(* IEC 61131-3 sources: plc-st-coding-agent/progress/evidence/f14_v5_public_pilot_20261112/jobs/custom_minimax-m27, 20 files *)

(* ---- public-easy-01.candidate_01.st ---- *)
FUNCTION_BLOCK FillingLineControl
VAR_INPUT
    bottleSensor          : BOOL;
    cleaningConfirmButton : BOOL;
    fillingConfirmButton  : BOOL;
    cappingConfirmButton  : BOOL;
    packingConfirmButton  : BOOL;
    finishedButton        : BOOL;
END_VAR
VAR_OUTPUT
    Pump_Motor       : BOOL;
    Filling_Valve    : BOOL;
    Capping_Machine  : BOOL;
    Packing_Machine  : BOOL;
    Completion_Light : BOOL;
END_VAR
VAR
    eState : INT;
END_VAR

// ENGINEERING_CONTRACT
// States: 0=IDLE, 1=CLEANING, 2=FILLING, 3=CAPPING, 4=PACKING, 5=COMPLETED
// PUB003: bottleSensor triggers pump motor continuously (retriggers if bottle stays)
// PUB004-PUB007: Each confirm button advances to next stage; next output activates immediately
// PUB008: finishedButton resets to IDLE; all outputs deactivate, Completion_Light clears
// Output retention: No output holds state beyond its stage; Completion_Light is latched until reset
// Same-scan priority: Transition logic evaluated after output assignments per state
// Boundaries: bottleSensor edge-sensitive to detected; confirm buttons level-triggered per stage

CASE eState OF
    0: // IDLE
        Pump_Motor       := FALSE;
        Filling_Valve    := FALSE;
        Capping_Machine  := FALSE;
        Packing_Machine  := FALSE;
        Completion_Light := FALSE;
        IF bottleSensor THEN
            eState := 1;
        END_IF;

    1: // CLEANING
        Pump_Motor       := TRUE;
        Filling_Valve    := FALSE;
        Capping_Machine  := FALSE;
        Packing_Machine  := FALSE;
        Completion_Light := FALSE;
        IF cleaningConfirmButton THEN
            eState := 2;
        END_IF;

    2: // FILLING
        Pump_Motor       := FALSE;
        Filling_Valve    := TRUE;
        Capping_Machine  := FALSE;
        Packing_Machine  := FALSE;
        Completion_Light := FALSE;
        IF fillingConfirmButton THEN
            eState := 3;
        END_IF;

    3: // CAPPING
        Pump_Motor       := FALSE;
        Filling_Valve    := FALSE;
        Capping_Machine  := TRUE;
        Packing_Machine  := FALSE;
        Completion_Light := FALSE;
        IF cappingConfirmButton THEN
            eState := 4;
        END_IF;

    4: // PACKING
        Pump_Motor       := FALSE;
        Filling_Valve    := FALSE;
        Capping_Machine  := FALSE;
        Packing_Machine  := TRUE;
        Completion_Light := FALSE;
        IF packingConfirmButton THEN
            eState := 5;
        END_IF;

    5: // COMPLETED
        Pump_Motor       := FALSE;
        Filling_Valve    := FALSE;
        Capping_Machine  := FALSE;
        Packing_Machine  := FALSE;
        Completion_Light := TRUE;
        IF finishedButton THEN
            eState := 0;
        END_IF;

END_CASE;

END_FUNCTION_BLOCK

(* ---- public-easy-01.candidate_02.st ---- *)
FUNCTION_BLOCK FillingLineControl
VAR_INPUT
    bottleSensor          : BOOL;
    cleaningConfirmButton : BOOL;
    fillingConfirmButton  : BOOL;
    cappingConfirmButton  : BOOL;
    packingConfirmButton  : BOOL;
    finishedButton        : BOOL;
END_VAR
VAR_OUTPUT
    Pump_Motor       : BOOL;
    Filling_Valve    : BOOL;
    Capping_Machine  : BOOL;
    Packing_Machine  : BOOL;
    Completion_Light : BOOL;
END_VAR
VAR
    eState    : INT;
    nextState : INT;
END_VAR

// ENGINEERING_CONTRACT
// States: 0=IDLE, 1=CLEANING, 2=FILLING, 3=CAPPING, 4=PACKING, 5=COMPLETED
// PUB003: bottleSensor triggers pump motor continuously (retriggers if bottle stays)
// PUB004-PUB007: Each confirm button advances to next stage; next output activates immediately
// PUB008: finishedButton resets to IDLE; all outputs deactivate, Completion_Light clears
// Output retention: No output holds state beyond its stage; Completion_Light is latched until reset
// Same-scan priority: Two-CASE pattern prevents premature output assignment during transition evaluation
// Boundaries: bottleSensor edge-sensitive to detected; confirm buttons level-triggered per stage

nextState := eState;
CASE eState OF
    0:
        IF bottleSensor THEN
            nextState := 1;
        END_IF;
    1:
        IF cleaningConfirmButton THEN
            nextState := 2;
        END_IF;
    2:
        IF fillingConfirmButton THEN
            nextState := 3;
        END_IF;
    3:
        IF cappingConfirmButton THEN
            nextState := 4;
        END_IF;
    4:
        IF packingConfirmButton THEN
            nextState := 5;
        END_IF;
    5:
        IF finishedButton THEN
            nextState := 0;
        END_IF;
END_CASE;

eState := nextState;

CASE eState OF
    0:
        Pump_Motor       := FALSE;
        Filling_Valve    := FALSE;
        Capping_Machine  := FALSE;
        Packing_Machine  := FALSE;
        Completion_Light := FALSE;
    1:
        Pump_Motor       := TRUE;
        Filling_Valve    := FALSE;
        Capping_Machine  := FALSE;
        Packing_Machine  := FALSE;
        Completion_Light := FALSE;
    2:
        Pump_Motor       := FALSE;
        Filling_Valve    := TRUE;
        Capping_Machine  := FALSE;
        Packing_Machine  := FALSE;
        Completion_Light := FALSE;
    3:
        Pump_Motor       := FALSE;
        Filling_Valve    := FALSE;
        Capping_Machine  := TRUE;
        Packing_Machine  := FALSE;
        Completion_Light := FALSE;
    4:
        Pump_Motor       := FALSE;
        Filling_Valve    := FALSE;
        Capping_Machine  := FALSE;
        Packing_Machine  := TRUE;
        Completion_Light := FALSE;
    5:
        Pump_Motor       := FALSE;
        Filling_Valve    := FALSE;
        Capping_Machine  := FALSE;
        Packing_Machine  := FALSE;
        Completion_Light := TRUE;
END_CASE;

END_FUNCTION_BLOCK

(* ---- public-easy-01.raw_candidate_01.st ---- *)
FUNCTION_BLOCK FillingLineControl
VAR_INPUT
    bottleSensor          : BOOL;
    cleaningConfirmButton : BOOL;
    fillingConfirmButton  : BOOL;
    cappingConfirmButton  : BOOL;
    packingConfirmButton  : BOOL;
    finishedButton        : BOOL;
END_VAR
VAR_OUTPUT
    Pump_Motor       : BOOL;
    Filling_Valve    : BOOL;
    Capping_Machine  : BOOL;
    Packing_Machine  : BOOL;
    Completion_Light : BOOL;
END_VAR
VAR
    eState : INT;
END_VAR

// ENGINEERING_CONTRACT
// States: 0=IDLE, 1=CLEANING, 2=FILLING, 3=CAPPING, 4=PACKING, 5=COMPLETED
// PUB003: bottleSensor triggers pump motor continuously (retriggers if bottle stays)
// PUB004-PUB007: Each confirm button advances to next stage; next output activates immediately
// PUB008: finishedButton resets to IDLE; all outputs deactivate, Completion_Light clears
// Output retention: No output holds state beyond its stage; Completion_Light is latched until reset
// Same-scan priority: Transition logic evaluated after output assignments per state
// Boundaries: bottleSensor edge-sensitive to detected; confirm buttons level-triggered per stage

CASE eState OF
    0: // IDLE
        Pump_Motor       := FALSE;
        Filling_Valve    := FALSE;
        Capping_Machine  := FALSE;
        Packing_Machine  := FALSE;
        Completion_Light := FALSE;
        IF bottleSensor THEN
            eState := 1;
        END_IF

    1: // CLEANING
        Pump_Motor       := TRUE;
        Filling_Valve    := FALSE;
        Capping_Machine  := FALSE;
        Packing_Machine  := FALSE;
        Completion_Light := FALSE;
        IF cleaningConfirmButton THEN
            eState := 2;
        END_IF

    2: // FILLING
        Pump_Motor       := FALSE;
        Filling_Valve    := TRUE;
        Capping_Machine  := FALSE;
        Packing_Machine  := FALSE;
        Completion_Light := FALSE;
        IF fillingConfirmButton THEN
            eState := 3;
        END_IF

    3: // CAPPING
        Pump_Motor       := FALSE;
        Filling_Valve    := FALSE;
        Capping_Machine  := TRUE;
        Packing_Machine  := FALSE;
        Completion_Light := FALSE;
        IF cappingConfirmButton THEN
            eState := 4;
        END_IF

    4: // PACKING
        Pump_Motor       := FALSE;
        Filling_Valve    := FALSE;
        Capping_Machine  := FALSE;
        Packing_Machine  := TRUE;
        Completion_Light := FALSE;
        IF packingConfirmButton THEN
            eState := 5;
        END_IF

    5: // COMPLETED
        Pump_Motor       := FALSE;
        Filling_Valve    := FALSE;
        Capping_Machine  := FALSE;
        Packing_Machine  := FALSE;
        Completion_Light := TRUE;
        IF finishedButton THEN
            eState := 0;
        END_IF

END_CASE

END_FUNCTION_BLOCK

(* ---- public-easy-01.raw_candidate_02.st ---- *)
FUNCTION_BLOCK FillingLineControl
VAR_INPUT
    bottleSensor          : BOOL;
    cleaningConfirmButton : BOOL;
    fillingConfirmButton  : BOOL;
    cappingConfirmButton  : BOOL;
    packingConfirmButton  : BOOL;
    finishedButton        : BOOL;
END_VAR
VAR_OUTPUT
    Pump_Motor       : BOOL;
    Filling_Valve    : BOOL;
    Capping_Machine  : BOOL;
    Packing_Machine  : BOOL;
    Completion_Light : BOOL;
END_VAR
VAR
    eState    : INT;
    nextState : INT;
END_VAR

// ENGINEERING_CONTRACT
// States: 0=IDLE, 1=CLEANING, 2=FILLING, 3=CAPPING, 4=PACKING, 5=COMPLETED
// PUB003: bottleSensor triggers pump motor continuously (retriggers if bottle stays)
// PUB004-PUB007: Each confirm button advances to next stage; next output activates immediately
// PUB008: finishedButton resets to IDLE; all outputs deactivate, Completion_Light clears
// Output retention: No output holds state beyond its stage; Completion_Light is latched until reset
// Same-scan priority: Two-CASE pattern prevents premature output assignment during transition evaluation
// Boundaries: bottleSensor edge-sensitive to detected; confirm buttons level-triggered per stage

nextState := eState;
CASE eState OF
    0:
        IF bottleSensor THEN
            nextState := 1;
        END_IF;
    1:
        IF cleaningConfirmButton THEN
            nextState := 2;
        END_IF;
    2:
        IF fillingConfirmButton THEN
            nextState := 3;
        END_IF;
    3:
        IF cappingConfirmButton THEN
            nextState := 4;
        END_IF;
    4:
        IF packingConfirmButton THEN
            nextState := 5;
        END_IF;
    5:
        IF finishedButton THEN
            nextState := 0;
        END_IF;
END_CASE;

eState := nextState;

CASE eState OF
    0:
        Pump_Motor       := FALSE;
        Filling_Valve    := FALSE;
        Capping_Machine  := FALSE;
        Packing_Machine  := FALSE;
        Completion_Light := FALSE;
    1:
        Pump_Motor       := TRUE;
        Filling_Valve    := FALSE;
        Capping_Machine  := FALSE;
        Packing_Machine  := FALSE;
        Completion_Light := FALSE;
    2:
        Pump_Motor       := FALSE;
        Filling_Valve    := TRUE;
        Capping_Machine  := FALSE;
        Packing_Machine  := FALSE;
        Completion_Light := FALSE;
    3:
        Pump_Motor       := FALSE;
        Filling_Valve    := FALSE;
        Capping_Machine  := TRUE;
        Packing_Machine  := FALSE;
        Completion_Light := FALSE;
    4:
        Pump_Motor       := FALSE;
        Filling_Valve    := FALSE;
        Capping_Machine  := FALSE;
        Packing_Machine  := TRUE;
        Completion_Light := FALSE;
    5:
        Pump_Motor       := FALSE;
        Filling_Valve    := FALSE;
        Capping_Machine  := FALSE;
        Packing_Machine  := FALSE;
        Completion_Light := TRUE;
END_CASE;

END_FUNCTION_BLOCK

(* ---- public-easy-04.candidate_01.st ---- *)
FUNCTION_BLOCK FB_JamPumpControl
VAR_INPUT
    VISCOSITY_OK    : BOOL;
    PASTE_E_STOP_NC : BOOL;
    DebounceTime    : TIME;
    CycleTime       : TIME;
END_VAR
VAR_OUTPUT
    VFD_RUN          : BOOL;
    PUMP_MAINT_DUE   : BOOL;
    PUMP_RUNTIME_ACC : LTIME;
END_VAR
VAR
    DebounceTimer : TON;
END_VAR

(*
ENGINEERING_CONTRACT - FB_JamPumpControl
================================================================================
| Output/State      | Activation           | Retention      | Reset/Deactivation           | Same-Scan | Units/Boundaries     |
|-------------------|----------------------|----------------|------------------------------|-----------|----------------------|
| VFD_RUN           | ESTOP AND vis_valid  | Hold TRUE      | Immediate: ESTOP=FALSE or    | ESTOP pri | Boolean              |
|                   |                      |                | viscosity_valid=FALSE        |           |                      |
| viscosity_valid   | DebounceTimer.Q=TRUE | Hold TRUE      | Immediate on VISCOSITY_OK=   | -         | Internal TON state   |
|                   |                      |                | FALSE or PASTE_E_STOP_NC=FALSE|          |                      |
| PUMP_RUNTIME_ACC  | Add CycleTime when   | Retain when    | Power-up init to 0 LTIME     | -         | LTIME (nanoseconds)  |
|                   | VFD_RUN=TRUE         | VFD_RUN=FALSE  |                              |           |                      |
| PUMP_MAINT_DUE    | ACC >= 500h (1.8e12ns)| Indefinite    | None (informational only)    | -         | Boolean              |
================================================================================
PUB001: Jam transfer pump control with viscosity debouncing, E-stop priority.
PUB002: VISCOSITY_OK debounced after DebounceTime; invalidated immediately on FALSE.
PUB003: VFD_RUN requires PASTE_E_STOP_NC=TRUE AND viscosity_valid; E-stop clears debounce.
PUB004: PUMP_RUNTIME_ACC accumulates via CycleTime only when VFD_RUN=TRUE; retains.
PUB005: PUMP_MAINT_DUE at 500h; informational, non-interlocking.
PUB006: Power-up: VFD_RUN=FALSE, PUMP_RUNTIME_ACC=0, PUMP_MAINT_DUE=FALSE.
================================================================================
*)

// Debounce viscosity signal
// Start timer when viscosity good AND E-stop permits; reset on E-stop loss or viscosity drop
DebounceTimer(
    IN  := VISCOSITY_OK AND PASTE_E_STOP_NC,
    PT  := DebounceTime
);

// Pump runs only when E-stop is active AND viscosity has been continuously valid for DebounceTime
VFD_RUN := PASTE_E_STOP_NC AND DebounceTimer.Q;

// Accumulate runtime while pump is running
IF VFD_RUN THEN
    PUMP_RUNTIME_ACC := PUMP_RUNTIME_ACC + LTIME_TO_LTIME(CycleTime);
END_IF;

// Maintenance due indication at 500 hours (500 * 3600 * 1000 * 1000000 nanoseconds)
PUMP_MAINT_DUE := (PUMP_RUNTIME_ACC >= T#500h) OR PUMP_MAINT_DUE;

END_FUNCTION_BLOCK

(* ---- public-easy-04.candidate_02.st ---- *)
FUNCTION_BLOCK FB_JamPumpControl
VAR_INPUT
    VISCOSITY_OK    : BOOL;
    PASTE_E_STOP_NC : BOOL;
    DebounceTime    : TIME;
    CycleTime       : TIME;
END_VAR
VAR_OUTPUT
    VFD_RUN          : BOOL;
    PUMP_MAINT_DUE   : BOOL;
    PUMP_RUNTIME_ACC : LTIME;
END_VAR
VAR
    DebounceTimer : TON;
END_VAR

(*
ENGINEERING_CONTRACT - FB_JamPumpControl
================================================================================
| Output/State      | Activation           | Retention      | Reset/Deactivation           | Same-Scan | Units/Boundaries     |
|-------------------|----------------------|----------------|------------------------------|-----------|----------------------|
| VFD_RUN           | ESTOP AND vis_valid  | Hold TRUE      | Immediate: ESTOP=FALSE or    | ESTOP pri | Boolean              |
|                   |                      |                | viscosity_valid=FALSE        |           |                      |
| viscosity_valid   | DebounceTimer.Q=TRUE | Hold TRUE      | Immediate on VISCOSITY_OK=   | -         | Internal TON state   |
|                   |                      |                | FALSE or PASTE_E_STOP_NC=FALSE|          |                      |
| PUMP_RUNTIME_ACC  | Add CycleTime when   | Retain when    | Power-up init to 0 LTIME     | -         | LTIME (nanoseconds)  |
|                   | VFD_RUN=TRUE         | VFD_RUN=FALSE  |                              |           |                      |
| PUMP_MAINT_DUE    | ACC >= 500h          | Indefinite    | None (informational only)    | -         | Boolean              |
================================================================================
PUB001: Jam transfer pump control with viscosity debouncing, E-stop priority.
PUB002: VISCOSITY_OK debounced after DebounceTime; invalidated immediately on FALSE.
PUB003: VFD_RUN requires PASTE_E_STOP_NC=TRUE AND viscosity_valid; E-stop clears debounce.
PUB004: PUMP_RUNTIME_ACC accumulates via CycleTime only when VFD_RUN=TRUE; retains.
PUB005: PUMP_MAINT_DUE at 500h; informational, non-interlocking.
PUB006: Power-up: VFD_RUN=FALSE, PUMP_RUNTIME_ACC=0, PUMP_MAINT_DUE=FALSE.
================================================================================
*)

// Debounce viscosity signal
// TON.IN resets (ET=0) immediately when PASTE_E_STOP_NC or VISCOSITY_OK goes FALSE
DebounceTimer(
    IN := VISCOSITY_OK AND PASTE_E_STOP_NC,
    PT := DebounceTime
);

// Pump runs only when E-stop is active AND viscosity has been continuously valid for DebounceTime
VFD_RUN := PASTE_E_STOP_NC AND DebounceTimer.Q;

// Accumulate runtime while pump is running
IF VFD_RUN THEN
    PUMP_RUNTIME_ACC := PUMP_RUNTIME_ACC + TIME_TO_LTIME(CycleTime);
END_IF;

// Maintenance due indication at 500 hours
PUMP_MAINT_DUE := PUMP_RUNTIME_ACC >= LTIME#500h;

END_FUNCTION_BLOCK

(* ---- public-easy-04.raw_candidate_01.st ---- *)
FUNCTION_BLOCK FB_JamPumpControl
VAR_INPUT
    VISCOSITY_OK    : BOOL;
    PASTE_E_STOP_NC : BOOL;
    DebounceTime    : TIME;
    CycleTime       : TIME;
END_VAR
VAR_OUTPUT
    VFD_RUN          : BOOL;
    PUMP_MAINT_DUE   : BOOL;
    PUMP_RUNTIME_ACC : LTIME;
END_VAR
VAR
    DebounceTimer : TON;
END_VAR

(*
ENGINEERING_CONTRACT - FB_JamPumpControl
================================================================================
| Output/State      | Activation           | Retention      | Reset/Deactivation           | Same-Scan | Units/Boundaries     |
|-------------------|----------------------|----------------|------------------------------|-----------|----------------------|
| VFD_RUN           | ESTOP AND vis_valid  | Hold TRUE      | Immediate: ESTOP=FALSE or    | ESTOP pri | Boolean              |
|                   |                      |                | viscosity_valid=FALSE        |           |                      |
| viscosity_valid   | DebounceTimer.Q=TRUE | Hold TRUE      | Immediate on VISCOSITY_OK=   | -         | Internal TON state   |
|                   |                      |                | FALSE or PASTE_E_STOP_NC=FALSE|          |                      |
| PUMP_RUNTIME_ACC  | Add CycleTime when   | Retain when    | Power-up init to 0 LTIME     | -         | LTIME (nanoseconds)  |
|                   | VFD_RUN=TRUE         | VFD_RUN=FALSE  |                              |           |                      |
| PUMP_MAINT_DUE    | ACC >= 500h (1.8e12ns)| Indefinite    | None (informational only)    | -         | Boolean              |
================================================================================
PUB001: Jam transfer pump control with viscosity debouncing, E-stop priority.
PUB002: VISCOSITY_OK debounced after DebounceTime; invalidated immediately on FALSE.
PUB003: VFD_RUN requires PASTE_E_STOP_NC=TRUE AND viscosity_valid; E-stop clears debounce.
PUB004: PUMP_RUNTIME_ACC accumulates via CycleTime only when VFD_RUN=TRUE; retains.
PUB005: PUMP_MAINT_DUE at 500h; informational, non-interlocking.
PUB006: Power-up: VFD_RUN=FALSE, PUMP_RUNTIME_ACC=0, PUMP_MAINT_DUE=FALSE.
================================================================================
*)

// Debounce viscosity signal
// Start timer when viscosity good AND E-stop permits; reset on E-stop loss or viscosity drop
DebounceTimer(
    IN  := VISCOSITY_OK AND PASTE_E_STOP_NC,
    PT  := DebounceTime
);

// Pump runs only when E-stop is active AND viscosity has been continuously valid for DebounceTime
VFD_RUN := PASTE_E_STOP_NC AND DebounceTimer.Q;

// Accumulate runtime while pump is running
IF VFD_RUN THEN
    PUMP_RUNTIME_ACC := PUMP_RUNTIME_ACC + LTIME_TO_LTIME(CycleTime);
END_IF

// Maintenance due indication at 500 hours (500 * 3600 * 1000 * 1000000 nanoseconds)
PUMP_MAINT_DUE := (PUMP_RUNTIME_ACC >= T#500h) OR PUMP_MAINT_DUE;

END_FUNCTION_BLOCK

(* ---- public-easy-04.raw_candidate_02.st ---- *)
FUNCTION_BLOCK FB_JamPumpControl
VAR_INPUT
    VISCOSITY_OK    : BOOL;
    PASTE_E_STOP_NC : BOOL;
    DebounceTime    : TIME;
    CycleTime       : TIME;
END_VAR
VAR_OUTPUT
    VFD_RUN          : BOOL;
    PUMP_MAINT_DUE   : BOOL;
    PUMP_RUNTIME_ACC : LTIME;
END_VAR
VAR
    DebounceTimer : TON;
END_VAR

(*
ENGINEERING_CONTRACT - FB_JamPumpControl
================================================================================
| Output/State      | Activation           | Retention      | Reset/Deactivation           | Same-Scan | Units/Boundaries     |
|-------------------|----------------------|----------------|------------------------------|-----------|----------------------|
| VFD_RUN           | ESTOP AND vis_valid  | Hold TRUE      | Immediate: ESTOP=FALSE or    | ESTOP pri | Boolean              |
|                   |                      |                | viscosity_valid=FALSE        |           |                      |
| viscosity_valid   | DebounceTimer.Q=TRUE | Hold TRUE      | Immediate on VISCOSITY_OK=   | -         | Internal TON state   |
|                   |                      |                | FALSE or PASTE_E_STOP_NC=FALSE|          |                      |
| PUMP_RUNTIME_ACC  | Add CycleTime when   | Retain when    | Power-up init to 0 LTIME     | -         | LTIME (nanoseconds)  |
|                   | VFD_RUN=TRUE         | VFD_RUN=FALSE  |                              |           |                      |
| PUMP_MAINT_DUE    | ACC >= 500h          | Indefinite    | None (informational only)    | -         | Boolean              |
================================================================================
PUB001: Jam transfer pump control with viscosity debouncing, E-stop priority.
PUB002: VISCOSITY_OK debounced after DebounceTime; invalidated immediately on FALSE.
PUB003: VFD_RUN requires PASTE_E_STOP_NC=TRUE AND viscosity_valid; E-stop clears debounce.
PUB004: PUMP_RUNTIME_ACC accumulates via CycleTime only when VFD_RUN=TRUE; retains.
PUB005: PUMP_MAINT_DUE at 500h; informational, non-interlocking.
PUB006: Power-up: VFD_RUN=FALSE, PUMP_RUNTIME_ACC=0, PUMP_MAINT_DUE=FALSE.
================================================================================
*)

// Debounce viscosity signal
// TON.IN resets (ET=0) immediately when PASTE_E_STOP_NC or VISCOSITY_OK goes FALSE
DebounceTimer(
    IN := VISCOSITY_OK AND PASTE_E_STOP_NC,
    PT := DebounceTime
);

// Pump runs only when E-stop is active AND viscosity has been continuously valid for DebounceTime
VFD_RUN := PASTE_E_STOP_NC AND DebounceTimer.Q;

// Accumulate runtime while pump is running
IF VFD_RUN THEN
    PUMP_RUNTIME_ACC := PUMP_RUNTIME_ACC + TIME_TO_LTIME(CycleTime);
END_IF;

// Maintenance due indication at 500 hours
PUMP_MAINT_DUE := PUMP_RUNTIME_ACC >= LTIME#500h;

END_FUNCTION_BLOCK

(* ---- public-hard-03.candidate_01.st ---- *)
FUNCTION_BLOCK FB_RecipeManagement
VAR_INPUT
    addRecipe     : BOOL;
    deleteRecipe  : BOOL;
    modifyRecipe  : BOOL;
    queryRecipe   : BOOL;
    recipeIn      : ST_Recipe;
END_VAR
VAR_OUTPUT
    recipeAdded       : BOOL;
    recipeDeleted     : BOOL;
    recipeModified    : BOOL;
    recipeQueryResult : ST_Recipe;
    error             : BOOL;
    status            : WORD;
END_VAR
VAR_IN_OUT
    recipe : ARRAY[1..10] OF ST_Recipe;
END_VAR
VAR
    fbAddR    : R_TRIG;
    fbDeleteR : R_TRIG;
    fbModifyR : R_TRIG;
    fbQueryR  : R_TRIG;
    idx       : INT;
    foundIdx  : INT;
    emptyIdx  : INT;
    hasFound  : BOOL;
    hasEmpty  : BOOL;
END_VAR

(* ENGINEERING_CONTRACT
| Output/State       | Activation           | Retention     | Reset/Deactivation           | Same-scan Priority | Units/Boundaries              |
|--------------------|----------------------|---------------|------------------------------|--------------------|-------------------------------|
| recipeAdded        | addRecipe rising edge| FALSE 1 scan  | Auto-clear next scan         | Highest            | BOOL                          |
| recipeDeleted      | deleteRecipe rising  | FALSE 1 scan  | Auto-clear next scan         | Highest            | BOOL                          |
| recipeModified     | modifyRecipe rising  | FALSE 1 scan  | Auto-clear next scan         | Highest            | BOOL                          |
| recipeQueryResult  | queryRecipe success  | Held          | Cleared on next query        | -                  | ST_Recipe                     |
| error              | Any operation fails  | Held          | Cleared on next success      | -                  | BOOL                          |
| status             | Set on error/success | Held          | 16#0000 on success           | -                  | WORD: 16#0000,16#8001-16#8005 |
PUB: PUB001,PUB002,PUB003,PUB004,PUB005,PUB006,PUB008,PUB009,PUB010,PUB011,PUB012
*)
BEGIN
    // Rising edge detection for all trigger inputs
    fbAddR(CLK := addRecipe);
    fbDeleteR(CLK := deleteRecipe);
    fbModifyR(CLK := modifyRecipe);
    fbQueryR(CLK := queryRecipe);

    // Default: clear success outputs each scan (latched for one scan then auto-reset)
    recipeAdded   := FALSE;
    recipeDeleted := FALSE;
    recipeModified:= FALSE;

    // QUERY operation (PUB006, PUB009, PUB012)
    IF fbQueryR.Q THEN
        hasFound := FALSE;
        foundIdx := 0;
        FOR idx := 1 TO 10 DO
            IF recipe[idx].recipeID = recipeIn.recipeID AND recipeIn.recipeID <> 0 THEN
                hasFound := TRUE;
                foundIdx := idx;
                EXIT;
            END_IF;
        END_FOR;

        IF hasFound THEN
            recipeQueryResult := recipe[foundIdx];
            error   := FALSE;
            status  := 16#0000;
        ELSE
            // Clear query result when not found
            recipeQueryResult.recipeID            := 0;
            recipeQueryResult.ingredientType      := 0;
            recipeQueryResult.ingredientRatio     := 0.0;
            recipeQueryResult.productionTemperature := 0.0;
            error   := TRUE;
            status  := 16#8001; // Recipe not found
        END_IF;
    END_IF;

    // ADD operation (PUB004, PUB008, PUB010)
    IF fbAddR.Q THEN
        hasFound := FALSE;
        hasEmpty := FALSE;
        emptyIdx := 0;
        foundIdx := 0;

        FOR idx := 1 TO 10 DO
            IF recipe[idx].recipeID = recipeIn.recipeID AND recipeIn.recipeID <> 0 THEN
                hasFound := TRUE;
                foundIdx := idx;
                EXIT;
            END_IF;
        END_FOR;

        IF NOT hasFound THEN
            FOR idx := 1 TO 10 DO
                IF recipe[idx].recipeID = 0 THEN
                    hasEmpty := TRUE;
                    emptyIdx := idx;
                    EXIT;
                END_IF;
            END_FOR;
        END_IF;

        IF hasFound THEN
            error  := TRUE;
            status := 16#8002; // Duplicate recipe ID
        ELSIF NOT hasEmpty THEN
            error  := TRUE;
            status := 16#8003; // No empty slot
        ELSE
            // Store in smallest-index empty slot (PUB010)
            recipe[emptyIdx] := recipeIn;
            recipeAdded      := TRUE;
            error            := FALSE;
            status           := 16#0000;
        END_IF;
    END_IF;

    // DELETE operation (PUB005, PUB008, PUB011)
    IF fbDeleteR.Q THEN
        hasFound := FALSE;
        foundIdx := 0;

        FOR idx := 1 TO 10 DO
            IF recipe[idx].recipeID = recipeIn.recipeID AND recipeIn.recipeID <> 0 THEN
                hasFound := TRUE;
                foundIdx := idx;
                EXIT;
            END_IF;
        END_FOR;

        IF hasFound THEN
            // Set recipeID to 0 to mark as empty slot (PUB011)
            recipe[foundIdx].recipeID := 0;
            recipeDeleted             := TRUE;
            error                     := FALSE;
            status                    := 16#0000;
        ELSE
            error  := TRUE;
            status := 16#8004; // Recipe not found
        END_IF;
    END_IF;

    // MODIFY operation (PUB005, PUB008, PUB012)
    IF fbModifyR.Q THEN
        hasFound := FALSE;
        foundIdx := 0;

        FOR idx := 1 TO 10 DO
            IF recipe[idx].recipeID = recipeIn.recipeID AND recipeIn.recipeID <> 0 THEN
                hasFound := TRUE;
                foundIdx := idx;
                EXIT;
            END_IF;
        END_FOR;

        IF hasFound THEN
            // Replace existing recipe with input recipe (PUB012)
            recipe[foundIdx] := recipeIn;
            recipeModified   := TRUE;
            error            := FALSE;
            status           := 16#0000;
        ELSE
            error  := TRUE;
            status := 16#8005; // Recipe not found
        END_IF;
    END_IF;
END_FUNCTION_BLOCK

(* ---- public-hard-03.candidate_02.st ---- *)
TYPE
    ST_Recipe : STRUCT
        recipeID             : INT;
        ingredientType       : INT;
        ingredientRatio      : REAL;
        productionTemperature: REAL;
    END_STRUCT
END_TYPE;

FUNCTION_BLOCK FB_RecipeManagement
VAR_INPUT
    addRecipe    : BOOL;
    deleteRecipe : BOOL;
    modifyRecipe : BOOL;
    queryRecipe  : BOOL;
    recipeIn     : ST_Recipe;
END_VAR
VAR_OUTPUT
    recipeAdded       : BOOL;
    recipeDeleted     : BOOL;
    recipeModified    : BOOL;
    recipeQueryResult : ST_Recipe;
    error             : BOOL;
    status            : WORD;
END_VAR
VAR_IN_OUT
    recipe : ARRAY[1..10] OF ST_Recipe;
END_VAR
VAR
    fbAddR    : R_TRIG;
    fbDeleteR : R_TRIG;
    fbModifyR : R_TRIG;
    fbQueryR  : R_TRIG;
    idx       : INT;
    foundIdx  : INT;
    emptyIdx  : INT;
    hasFound  : BOOL;
    hasEmpty  : BOOL;
END_VAR

(* ENGINEERING_CONTRACT
| Output/State       | Activation           | Retention     | Reset/Deactivation           | Same-scan Priority | Units/Boundaries              |
|--------------------|----------------------|---------------|------------------------------|--------------------|-------------------------------|
| recipeAdded        | addRecipe rising edge| FALSE 1 scan  | Auto-clear next scan         | Highest            | BOOL                          |
| recipeDeleted      | deleteRecipe rising  | FALSE 1 scan  | Auto-clear next scan         | Highest            | BOOL                          |
| recipeModified     | modifyRecipe rising  | FALSE 1 scan  | Auto-clear next scan         | Highest            | BOOL                          |
| recipeQueryResult  | queryRecipe success  | Held          | Cleared on next query        | -                  | ST_Recipe                     |
| error              | Any operation fails  | Held          | Cleared on next success      | -                  | BOOL                          |
| status             | Set on error/success | Held          | 16#0000 on success           | -                  | WORD: 16#0000,16#8001-16#8005 |
PUB: PUB001,PUB002,PUB003,PUB004,PUB005,PUB006,PUB008,PUB009,PUB010,PUB011,PUB012
*)
    fbAddR(CLK := addRecipe);
    fbDeleteR(CLK := deleteRecipe);
    fbModifyR(CLK := modifyRecipe);
    fbQueryR(CLK := queryRecipe);

    recipeAdded   := FALSE;
    recipeDeleted := FALSE;
    recipeModified:= FALSE;

    IF fbQueryR.Q THEN
        hasFound := FALSE;
        foundIdx := 0;
        FOR idx := 1 TO 10 DO
            IF recipe[idx].recipeID = recipeIn.recipeID AND recipeIn.recipeID <> 0 THEN
                hasFound := TRUE;
                foundIdx := idx;
                EXIT;
            END_IF;
        END_FOR;

        IF hasFound THEN
            recipeQueryResult := recipe[foundIdx];
            error  := FALSE;
            status := 16#0000;
        ELSE
            recipeQueryResult.recipeID             := 0;
            recipeQueryResult.ingredientType       := 0;
            recipeQueryResult.ingredientRatio      := 0.0;
            recipeQueryResult.productionTemperature:= 0.0;
            error  := TRUE;
            status := 16#8001;
        END_IF;
    END_IF;

    IF fbAddR.Q THEN
        hasFound := FALSE;
        hasEmpty := FALSE;
        emptyIdx := 0;
        foundIdx := 0;

        FOR idx := 1 TO 10 DO
            IF recipe[idx].recipeID = recipeIn.recipeID AND recipeIn.recipeID <> 0 THEN
                hasFound := TRUE;
                foundIdx := idx;
                EXIT;
            END_IF;
        END_FOR;

        IF NOT hasFound THEN
            FOR idx := 1 TO 10 DO
                IF recipe[idx].recipeID = 0 THEN
                    hasEmpty := TRUE;
                    emptyIdx := idx;
                    EXIT;
                END_IF;
            END_FOR;
        END_IF;

        IF hasFound THEN
            error  := TRUE;
            status := 16#8002;
        ELSIF NOT hasEmpty THEN
            error  := TRUE;
            status := 16#8003;
        ELSE
            recipe[emptyIdx] := recipeIn;
            recipeAdded      := TRUE;
            error            := FALSE;
            status           := 16#0000;
        END_IF;
    END_IF;

    IF fbDeleteR.Q THEN
        hasFound := FALSE;
        foundIdx := 0;

        FOR idx := 1 TO 10 DO
            IF recipe[idx].recipeID = recipeIn.recipeID AND recipeIn.recipeID <> 0 THEN
                hasFound := TRUE;
                foundIdx := idx;
                EXIT;
            END_IF;
        END_FOR;

        IF hasFound THEN
            recipe[foundIdx].recipeID := 0;
            recipeDeleted             := TRUE;
            error                     := FALSE;
            status                    := 16#0000;
        ELSE
            error  := TRUE;
            status := 16#8004;
        END_IF;
    END_IF;

    IF fbModifyR.Q THEN
        hasFound := FALSE;
        foundIdx := 0;

        FOR idx := 1 TO 10 DO
            IF recipe[idx].recipeID = recipeIn.recipeID AND recipeIn.recipeID <> 0 THEN
                hasFound := TRUE;
                foundIdx := idx;
                EXIT;
            END_IF;
        END_FOR;

        IF hasFound THEN
            recipe[foundIdx] := recipeIn;
            recipeModified   := TRUE;
            error            := FALSE;
            status           := 16#0000;
        ELSE
            error  := TRUE;
            status := 16#8005;
        END_IF;
    END_IF;
END_FUNCTION_BLOCK

(* ---- public-hard-03.raw_candidate_01.st ---- *)
FUNCTION_BLOCK FB_RecipeManagement
VAR_INPUT
    addRecipe     : BOOL;
    deleteRecipe  : BOOL;
    modifyRecipe  : BOOL;
    queryRecipe   : BOOL;
    recipeIn      : ST_Recipe;
END_VAR
VAR_OUTPUT
    recipeAdded       : BOOL;
    recipeDeleted     : BOOL;
    recipeModified    : BOOL;
    recipeQueryResult : ST_Recipe;
    error             : BOOL;
    status            : WORD;
END_VAR
VAR_IN_OUT
    recipe : ARRAY[1..10] OF ST_Recipe;
END_VAR
VAR
    fbAddR    : R_TRIG;
    fbDeleteR : R_TRIG;
    fbModifyR : R_TRIG;
    fbQueryR  : R_TRIG;
    idx       : INT;
    foundIdx  : INT;
    emptyIdx  : INT;
    hasFound  : BOOL;
    hasEmpty  : BOOL;
END_VAR

(* ENGINEERING_CONTRACT
| Output/State       | Activation           | Retention     | Reset/Deactivation           | Same-scan Priority | Units/Boundaries              |
|--------------------|----------------------|---------------|------------------------------|--------------------|-------------------------------|
| recipeAdded        | addRecipe rising edge| FALSE 1 scan  | Auto-clear next scan         | Highest            | BOOL                          |
| recipeDeleted      | deleteRecipe rising  | FALSE 1 scan  | Auto-clear next scan         | Highest            | BOOL                          |
| recipeModified     | modifyRecipe rising  | FALSE 1 scan  | Auto-clear next scan         | Highest            | BOOL                          |
| recipeQueryResult  | queryRecipe success  | Held          | Cleared on next query        | -                  | ST_Recipe                     |
| error              | Any operation fails  | Held          | Cleared on next success      | -                  | BOOL                          |
| status             | Set on error/success | Held          | 16#0000 on success           | -                  | WORD: 16#0000,16#8001-16#8005 |
PUB: PUB001,PUB002,PUB003,PUB004,PUB005,PUB006,PUB008,PUB009,PUB010,PUB011,PUB012
*)
BEGIN
    // Rising edge detection for all trigger inputs
    fbAddR(CLK := addRecipe);
    fbDeleteR(CLK := deleteRecipe);
    fbModifyR(CLK := modifyRecipe);
    fbQueryR(CLK := queryRecipe);

    // Default: clear success outputs each scan (latched for one scan then auto-reset)
    recipeAdded   := FALSE;
    recipeDeleted := FALSE;
    recipeModified:= FALSE;

    // QUERY operation (PUB006, PUB009, PUB012)
    IF fbQueryR.Q THEN
        hasFound := FALSE;
        foundIdx := 0;
        FOR idx := 1 TO 10 DO
            IF recipe[idx].recipeID = recipeIn.recipeID AND recipeIn.recipeID <> 0 THEN
                hasFound := TRUE;
                foundIdx := idx;
                EXIT;
            END_IF;
        END_FOR;

        IF hasFound THEN
            recipeQueryResult := recipe[foundIdx];
            error   := FALSE;
            status  := 16#0000;
        ELSE
            // Clear query result when not found
            recipeQueryResult.recipeID            := 0;
            recipeQueryResult.ingredientType      := 0;
            recipeQueryResult.ingredientRatio     := 0.0;
            recipeQueryResult.productionTemperature := 0.0;
            error   := TRUE;
            status  := 16#8001; // Recipe not found
        END_IF;
    END_IF;

    // ADD operation (PUB004, PUB008, PUB010)
    IF fbAddR.Q THEN
        hasFound := FALSE;
        hasEmpty := FALSE;
        emptyIdx := 0;
        foundIdx := 0;

        FOR idx := 1 TO 10 DO
            IF recipe[idx].recipeID = recipeIn.recipeID AND recipeIn.recipeID <> 0 THEN
                hasFound := TRUE;
                foundIdx := idx;
                EXIT;
            END_IF;
        END_FOR;

        IF NOT hasFound THEN
            FOR idx := 1 TO 10 DO
                IF recipe[idx].recipeID = 0 THEN
                    hasEmpty := TRUE;
                    emptyIdx := idx;
                    EXIT;
                END_IF;
            END_FOR;
        END_IF;

        IF hasFound THEN
            error  := TRUE;
            status := 16#8002; // Duplicate recipe ID
        ELSIF NOT hasEmpty THEN
            error  := TRUE;
            status := 16#8003; // No empty slot
        ELSE
            // Store in smallest-index empty slot (PUB010)
            recipe[emptyIdx] := recipeIn;
            recipeAdded      := TRUE;
            error            := FALSE;
            status           := 16#0000;
        END_IF;
    END_IF;

    // DELETE operation (PUB005, PUB008, PUB011)
    IF fbDeleteR.Q THEN
        hasFound := FALSE;
        foundIdx := 0;

        FOR idx := 1 TO 10 DO
            IF recipe[idx].recipeID = recipeIn.recipeID AND recipeIn.recipeID <> 0 THEN
                hasFound := TRUE;
                foundIdx := idx;
                EXIT;
            END_IF;
        END_FOR;

        IF hasFound THEN
            // Set recipeID to 0 to mark as empty slot (PUB011)
            recipe[foundIdx].recipeID := 0;
            recipeDeleted             := TRUE;
            error                     := FALSE;
            status                    := 16#0000;
        ELSE
            error  := TRUE;
            status := 16#8004; // Recipe not found
        END_IF;
    END_IF;

    // MODIFY operation (PUB005, PUB008, PUB012)
    IF fbModifyR.Q THEN
        hasFound := FALSE;
        foundIdx := 0;

        FOR idx := 1 TO 10 DO
            IF recipe[idx].recipeID = recipeIn.recipeID AND recipeIn.recipeID <> 0 THEN
                hasFound := TRUE;
                foundIdx := idx;
                EXIT;
            END_IF;
        END_FOR;

        IF hasFound THEN
            // Replace existing recipe with input recipe (PUB012)
            recipe[foundIdx] := recipeIn;
            recipeModified   := TRUE;
            error            := FALSE;
            status           := 16#0000;
        ELSE
            error  := TRUE;
            status := 16#8005; // Recipe not found
        END_IF;
    END_IF;
END_FUNCTION_BLOCK

(* ---- public-hard-03.raw_candidate_02.st ---- *)
TYPE
    ST_Recipe : STRUCT
        recipeID             : INT;
        ingredientType       : INT;
        ingredientRatio      : REAL;
        productionTemperature: REAL;
    END_STRUCT
END_TYPE

FUNCTION_BLOCK FB_RecipeManagement
VAR_INPUT
    addRecipe    : BOOL;
    deleteRecipe : BOOL;
    modifyRecipe : BOOL;
    queryRecipe  : BOOL;
    recipeIn     : ST_Recipe;
END_VAR
VAR_OUTPUT
    recipeAdded       : BOOL;
    recipeDeleted     : BOOL;
    recipeModified    : BOOL;
    recipeQueryResult : ST_Recipe;
    error             : BOOL;
    status            : WORD;
END_VAR
VAR_IN_OUT
    recipe : ARRAY[1..10] OF ST_Recipe;
END_VAR
VAR
    fbAddR    : R_TRIG;
    fbDeleteR : R_TRIG;
    fbModifyR : R_TRIG;
    fbQueryR  : R_TRIG;
    idx       : INT;
    foundIdx  : INT;
    emptyIdx  : INT;
    hasFound  : BOOL;
    hasEmpty  : BOOL;
END_VAR

(* ENGINEERING_CONTRACT
| Output/State       | Activation           | Retention     | Reset/Deactivation           | Same-scan Priority | Units/Boundaries              |
|--------------------|----------------------|---------------|------------------------------|--------------------|-------------------------------|
| recipeAdded        | addRecipe rising edge| FALSE 1 scan  | Auto-clear next scan         | Highest            | BOOL                          |
| recipeDeleted      | deleteRecipe rising  | FALSE 1 scan  | Auto-clear next scan         | Highest            | BOOL                          |
| recipeModified     | modifyRecipe rising  | FALSE 1 scan  | Auto-clear next scan         | Highest            | BOOL                          |
| recipeQueryResult  | queryRecipe success  | Held          | Cleared on next query        | -                  | ST_Recipe                     |
| error              | Any operation fails  | Held          | Cleared on next success      | -                  | BOOL                          |
| status             | Set on error/success | Held          | 16#0000 on success           | -                  | WORD: 16#0000,16#8001-16#8005 |
PUB: PUB001,PUB002,PUB003,PUB004,PUB005,PUB006,PUB008,PUB009,PUB010,PUB011,PUB012
*)
    fbAddR(CLK := addRecipe);
    fbDeleteR(CLK := deleteRecipe);
    fbModifyR(CLK := modifyRecipe);
    fbQueryR(CLK := queryRecipe);

    recipeAdded   := FALSE;
    recipeDeleted := FALSE;
    recipeModified:= FALSE;

    IF fbQueryR.Q THEN
        hasFound := FALSE;
        foundIdx := 0;
        FOR idx := 1 TO 10 DO
            IF recipe[idx].recipeID = recipeIn.recipeID AND recipeIn.recipeID <> 0 THEN
                hasFound := TRUE;
                foundIdx := idx;
                EXIT;
            END_IF;
        END_FOR;

        IF hasFound THEN
            recipeQueryResult := recipe[foundIdx];
            error  := FALSE;
            status := 16#0000;
        ELSE
            recipeQueryResult.recipeID             := 0;
            recipeQueryResult.ingredientType       := 0;
            recipeQueryResult.ingredientRatio      := 0.0;
            recipeQueryResult.productionTemperature:= 0.0;
            error  := TRUE;
            status := 16#8001;
        END_IF;
    END_IF;

    IF fbAddR.Q THEN
        hasFound := FALSE;
        hasEmpty := FALSE;
        emptyIdx := 0;
        foundIdx := 0;

        FOR idx := 1 TO 10 DO
            IF recipe[idx].recipeID = recipeIn.recipeID AND recipeIn.recipeID <> 0 THEN
                hasFound := TRUE;
                foundIdx := idx;
                EXIT;
            END_IF;
        END_FOR;

        IF NOT hasFound THEN
            FOR idx := 1 TO 10 DO
                IF recipe[idx].recipeID = 0 THEN
                    hasEmpty := TRUE;
                    emptyIdx := idx;
                    EXIT;
                END_IF;
            END_FOR;
        END_IF;

        IF hasFound THEN
            error  := TRUE;
            status := 16#8002;
        ELSIF NOT hasEmpty THEN
            error  := TRUE;
            status := 16#8003;
        ELSE
            recipe[emptyIdx] := recipeIn;
            recipeAdded      := TRUE;
            error            := FALSE;
            status           := 16#0000;
        END_IF;
    END_IF;

    IF fbDeleteR.Q THEN
        hasFound := FALSE;
        foundIdx := 0;

        FOR idx := 1 TO 10 DO
            IF recipe[idx].recipeID = recipeIn.recipeID AND recipeIn.recipeID <> 0 THEN
                hasFound := TRUE;
                foundIdx := idx;
                EXIT;
            END_IF;
        END_FOR;

        IF hasFound THEN
            recipe[foundIdx].recipeID := 0;
            recipeDeleted             := TRUE;
            error                     := FALSE;
            status                    := 16#0000;
        ELSE
            error  := TRUE;
            status := 16#8004;
        END_IF;
    END_IF;

    IF fbModifyR.Q THEN
        hasFound := FALSE;
        foundIdx := 0;

        FOR idx := 1 TO 10 DO
            IF recipe[idx].recipeID = recipeIn.recipeID AND recipeIn.recipeID <> 0 THEN
                hasFound := TRUE;
                foundIdx := idx;
                EXIT;
            END_IF;
        END_FOR;

        IF hasFound THEN
            recipe[foundIdx] := recipeIn;
            recipeModified   := TRUE;
            error            := FALSE;
            status           := 16#0000;
        ELSE
            error  := TRUE;
            status := 16#8005;
        END_IF;
    END_IF;
END_FUNCTION_BLOCK

(* ---- public-medium-03.candidate_01.st ---- *)
FUNCTION_BLOCK FB_MovingAverage
VAR_INPUT
    cyclicExecution : BOOL;
    trigger         : BOOL;
    value           : LREAL;
    windowSize      : INT;
    reset           : BOOL;
END_VAR

VAR_OUTPUT
    average         : LREAL;
    windowSizeReached: BOOL;
    error           : BOOL;
    status          : WORD;
END_VAR

VAR
    dataBuffer      : ARRAY[1..100] OF LREAL;
    currentIndex    : INT := 0;
    sampleCount     : INT := 0;
    sum             : LREAL := 0.0;
    lastTrigger     : BOOL := FALSE;
    lastWindowSize  : INT := 0;
END_VAR

(* =========================================================================
   ENGINEERING_CONTRACT - Moving Average Function Block

   PUB001: Moving arithmetic mean via FIFO sliding window
   PUB002: cyclicExecution TRUE -> auto-update every scan (no edge needed)
   PUB003: trigger rising edge -> single-sample update per edge
   PUB004: reset TRUE -> full state clear; windowSize validation 1..100

   OUTPUT BEHAVIOR TABLE:
   | Output            | Activation        | Retention    | Reset        | Units/Range          |
   |-------------------|-------------------|--------------|--------------|----------------------|
   | average           | on valid update   | holds last   | on reset     | LREAL, computed      |
   | windowSizeReached | when count == size| holds state  | on reset     | FALSE(0..n-1), TRUE(n)|
   | error             | windowSize !in[1,100]| holds    | on reset     | FALSE=ok, TRUE=error |
   | status            | 16#8200 on bad size| holds      | on reset     | 16#0000, 16#8200     |

   BOUNDARY/SAME-SCAN RULES:
   - windowSize change invalidates: reinit buffer, no error until next cycle
   - cyclicExecution dominates trigger; trigger ignored when cyclic=TRUE
   - Rising edge: lastTrigger (previous cycle) vs trigger (current)
   - Zero samples: average=0.0, windowSizeReached=FALSE
   - reset clears all state including error and status in same scan

   ========================================================================= *)

    // --- Reset handling (highest priority) ---
    IF reset THEN
        currentIndex     := 0;
        sampleCount      := 0;
        sum              := 0.0;
        average          := 0.0;
        windowSizeReached := FALSE;
        error            := FALSE;
        status           := 16#0000;
        lastTrigger      := FALSE;
        lastWindowSize   := 0;
        RETURN;
    END_IF;

    // --- Window size validation ---
    IF (windowSize < 1) OR (windowSize > 100) THEN
        error  := TRUE;
        status := 16#8200;
        RETURN;
    END_IF;

    // --- Reinitialize buffer when window size changes to valid value ---
    IF lastWindowSize <> windowSize THEN
        currentIndex     := 0;
        sampleCount      := 0;
        sum              := 0.0;
        average          := 0.0;
        windowSizeReached := FALSE;
        lastWindowSize   := windowSize;
    END_IF;

    // --- Execution trigger selection ---
    // PUB002: cyclicExecution TRUE -> update every scan
    // PUB003: trigger rising edge -> update per edge
    // Same-scan priority: cyclicExecution takes precedence
    IF cyclicExecution OR (trigger AND NOT lastTrigger) THEN
        // Advance circular buffer index
        currentIndex := (currentIndex MOD windowSize) + 1;

        // Subtract the value being overwritten from sum (FIFO principle)
        IF sampleCount >= windowSize THEN
            sum := sum - dataBuffer[currentIndex];
        END_IF;

        // Add new value to sum and buffer
        sum := sum + value;
        dataBuffer[currentIndex] := value;

        // Increment sample count up to window size
        IF sampleCount < windowSize THEN
            sampleCount := sampleCount + 1;
        END_IF;

        // Compute moving average (sum / current count)
        average := sum / TO_LREAL(sampleCount);

        // Update window reached flag
        windowSizeReached := (sampleCount >= windowSize);

        // Clear error on successful execution
        error  := FALSE;
        status := 16#0000;
    END_IF;

    // --- Latch last trigger state for edge detection ---
    lastTrigger := trigger;

END_FUNCTION_BLOCK

(* ---- public-medium-03.raw_candidate_01.st ---- *)
FUNCTION_BLOCK FB_MovingAverage
VAR_INPUT
    cyclicExecution : BOOL;
    trigger         : BOOL;
    value           : LREAL;
    windowSize      : INT;
    reset           : BOOL;
END_VAR

VAR_OUTPUT
    average         : LREAL;
    windowSizeReached: BOOL;
    error           : BOOL;
    status          : WORD;
END_VAR

VAR
    dataBuffer      : ARRAY[1..100] OF LREAL;
    currentIndex    : INT := 0;
    sampleCount     : INT := 0;
    sum             : LREAL := 0.0;
    lastTrigger     : BOOL := FALSE;
    lastWindowSize  : INT := 0;
END_VAR

(* =========================================================================
   ENGINEERING_CONTRACT - Moving Average Function Block

   PUB001: Moving arithmetic mean via FIFO sliding window
   PUB002: cyclicExecution TRUE -> auto-update every scan (no edge needed)
   PUB003: trigger rising edge -> single-sample update per edge
   PUB004: reset TRUE -> full state clear; windowSize validation 1..100

   OUTPUT BEHAVIOR TABLE:
   | Output            | Activation        | Retention    | Reset        | Units/Range          |
   |-------------------|-------------------|--------------|--------------|----------------------|
   | average           | on valid update   | holds last   | on reset     | LREAL, computed      |
   | windowSizeReached | when count == size| holds state  | on reset     | FALSE(0..n-1), TRUE(n)|
   | error             | windowSize !in[1,100]| holds    | on reset     | FALSE=ok, TRUE=error |
   | status            | 16#8200 on bad size| holds      | on reset     | 16#0000, 16#8200     |

   BOUNDARY/SAME-SCAN RULES:
   - windowSize change invalidates: reinit buffer, no error until next cycle
   - cyclicExecution dominates trigger; trigger ignored when cyclic=TRUE
   - Rising edge: lastTrigger (previous cycle) vs trigger (current)
   - Zero samples: average=0.0, windowSizeReached=FALSE
   - reset clears all state including error and status in same scan

   ========================================================================= *)

    // --- Reset handling (highest priority) ---
    IF reset THEN
        currentIndex     := 0;
        sampleCount      := 0;
        sum              := 0.0;
        average          := 0.0;
        windowSizeReached := FALSE;
        error            := FALSE;
        status           := 16#0000;
        lastTrigger      := FALSE;
        lastWindowSize   := 0;
        RETURN;
    END_IF

    // --- Window size validation ---
    IF (windowSize < 1) OR (windowSize > 100) THEN
        error  := TRUE;
        status := 16#8200;
        RETURN;
    END_IF

    // --- Reinitialize buffer when window size changes to valid value ---
    IF lastWindowSize <> windowSize THEN
        currentIndex     := 0;
        sampleCount      := 0;
        sum              := 0.0;
        average          := 0.0;
        windowSizeReached := FALSE;
        lastWindowSize   := windowSize;
    END_IF

    // --- Execution trigger selection ---
    // PUB002: cyclicExecution TRUE -> update every scan
    // PUB003: trigger rising edge -> update per edge
    // Same-scan priority: cyclicExecution takes precedence
    IF cyclicExecution OR (trigger AND NOT lastTrigger) THEN
        // Advance circular buffer index
        currentIndex := (currentIndex MOD windowSize) + 1;

        // Subtract the value being overwritten from sum (FIFO principle)
        IF sampleCount >= windowSize THEN
            sum := sum - dataBuffer[currentIndex];
        END_IF

        // Add new value to sum and buffer
        sum := sum + value;
        dataBuffer[currentIndex] := value;

        // Increment sample count up to window size
        IF sampleCount < windowSize THEN
            sampleCount := sampleCount + 1;
        END_IF

        // Compute moving average (sum / current count)
        average := sum / TO_LREAL(sampleCount);

        // Update window reached flag
        windowSizeReached := (sampleCount >= windowSize);

        // Clear error on successful execution
        error  := FALSE;
        status := 16#0000;
    END_IF

    // --- Latch last trigger state for edge detection ---
    lastTrigger := trigger;

END_FUNCTION_BLOCK

(* ---- public-medium-04.candidate_01.st ---- *)
FUNCTION_BLOCK FB_TemperatureControl
VAR_INPUT
    TemperatureSensorInput : REAL;
    SetTemperature         : REAL;
END_VAR
VAR_OUTPUT
    CurrentTemperature : REAL;
    SetTempDisplay     : REAL;
    HeaterStatus       : BOOL;
    OverheatProtection : BOOL;
    HeaterOutput       : BOOL;
END_VAR
VAR
    heaterOnTimer         : TON;
    overheatRecoveryTimer : TON;
    heaterOnTime          : LTIME := LTIME#5s;
    overheatWaitTime      : LTIME := LTIME#3s;
    overheatTriggered     : BOOL  := FALSE;
    sensorFault           : BOOL  := FALSE;
    heaterOnCondition     : BOOL  := FALSE;
    validTemperature      : REAL  := 0.0;
END_VAR
//---------------------------------------------------------------------------
// ENGINEERING_CONTRACT
// +-----------+-----------+-------------------------------+------+----------+
// | Output    | Activation| Retention/Reset               | Prior| Boundary |
// +-----------+-----------+-------------------------------+------+----------+
// | HeaterOut | Temp<Set  | Cleared on: fault, overheat,  | 1st  | PUB007   |
// |           | +no fault | temp>=Set (this scan),        |      | PUB003-5 |
// |           | +no OHP   | overheatTimer expired         |      |          |
// +-----------+-----------+-------------------------------+------+----------+
// | OverheatP | 5s heater | Reset after 3s recovery;      | 2nd  | PUB006   |
// |           | ON cont.  | cleared by overheatTimer.Q    |      |          |
// +-----------+-----------+-------------------------------+------+----------+
// | HeaterSt  | =HeaterOut| Same deactivation as above    | -    | PUB007   |
// +-----------+-----------+-------------------------------+------+----------+
// | CurrTemp  | Valid Rd  | Fault->0.0; else actual       | -    | PUB007   |
// +-----------+-----------+-------------------------------+------+----------+
// | SetTemp   | Always SetTemperature input               | -    | PUB007   |
// +-----------+-----------+-------------------------------+------+----------+
// | Sensor    | Input<0 OR >100 (edge-insensitive)       | Auto | PUB007   |
// | Fault     | Clears when input returns to [0..100]    | reset|          |
// +-----------+-----------+-------------------------------+------+----------+
// Same-scan priority order: Sensor Fault > Overheat > Temperature Comparison
// Timing: 5s continuous ON triggers OHP; 3s wait before OHP release
//---------------------------------------------------------------------------

    // PUB007: Sensor fault detection (outside [0,100])
    sensorFault := (TemperatureSensorInput < 0.0) OR (TemperatureSensorInput > 100.0);

    // PUB007: Display current temperature; show 0.0 on fault
    IF sensorFault THEN
        validTemperature := 0.0;
    ELSE
        validTemperature := TemperatureSensorInput;
    END_IF;

    // PUB003-PUB005: Temperature comparison
    // Heater request is TRUE when actual < set AND no fault
    heaterOnCondition := (TemperatureSensorInput < SetTemperature) AND NOT sensorFault;

    // PUB006: Heater-on accumulation timer
    heaterOnTimer(IN := heaterOnCondition AND NOT overheatTriggered, PT := heaterOnTime);

    // PUB006: Overheat trigger - ON > 5s
    IF heaterOnTimer.ET >= heaterOnTime AND NOT overheatTriggered THEN
        overheatTriggered := TRUE;
    END_IF;

    // PUB006: After overheat triggered, reset the accumulation timer so
    // ET returns to 0 while heater is suppressed; ON condition may still
    // be TRUE but the timer will be inactive until overheat clears.
    IF overheatTriggered THEN
        heaterOnTimer(IN := FALSE, PT := heaterOnTime);
    END_IF;

    // PUB006: Overheat recovery timer starts when overheatTriggered is TRUE
    // and runs for 3s; heaterOnCondition may still be TRUE during this wait.
    overheatRecoveryTimer(IN := overheatTriggered, PT := overheatWaitTime);

    // PUB006: Release overheat protection after 3s elapsed
    IF overheatRecoveryTimer.Q THEN
        overheatTriggered := FALSE;
    END_IF;

    // PUB007: Status outputs
    SetTempDisplay := SetTemperature;
    CurrentTemperature := validTemperature;
    HeaterStatus := heaterOnCondition AND NOT sensorFault AND NOT overheatTriggered;

    // PUB004/PUB005: HeaterOutput suppressed when sensor fault or overheat active
    HeaterOutput := heaterOnCondition AND NOT sensorFault AND NOT overheatTriggered;

END_FUNCTION_BLOCK

(* ---- public-medium-04.candidate_02.st ---- *)
FUNCTION_BLOCK FB_TemperatureControl
VAR_INPUT
    TemperatureSensorInput : REAL;
    SetTemperature         : REAL;
END_VAR
VAR_OUTPUT
    CurrentTemperature : REAL;
    SetTempDisplay     : REAL;
    HeaterStatus       : BOOL;
    OverheatProtection : BOOL;
    HeaterOutput       : BOOL;
END_VAR
VAR
    heaterOnTimer         : TON;
    overheatRecoveryTimer : TON;
    heaterOnTime          : TIME := TIME#5s;
    overheatWaitTime      : TIME := TIME#3s;
    overheatTriggered     : BOOL  := FALSE;
    sensorFault           : BOOL  := FALSE;
    heaterOnCondition     : BOOL  := FALSE;
    validTemperature      : REAL  := 0.0;
END_VAR
//---------------------------------------------------------------------------
// ENGINEERING_CONTRACT
// +-----------+-----------+-------------------------------+------+----------+
// | Output    | Activation| Retention/Reset               | Prior| Boundary |
// +-----------+-----------+-------------------------------+------+----------+
// | HeaterOut | Temp<Set  | Cleared on: fault, overheat,  | 1st  | PUB007   |
// |           | +no fault | temp>=Set (this scan),        |      | PUB003-5 |
// |           | +no OHP   | overheatTimer expired         |      |          |
// +-----------+-----------+-------------------------------+------+----------+
// | OverheatP | 5s heater | Reset after 3s recovery;      | 2nd  | PUB006   |
// |           | ON cont.  | cleared by overheatTimer.Q    |      |          |
// +-----------+-----------+-------------------------------+------+----------+
// | HeaterSt  | =HeaterOut| Same deactivation as above    | -    | PUB007   |
// +-----------+-----------+-------------------------------+------+----------+
// | CurrTemp  | Valid Rd  | Fault->0.0; else actual       | -    | PUB007   |
// +-----------+-----------+-------------------------------+------+----------+
// | SetTemp   | Always SetTemperature input               | -    | PUB007   |
// +-----------+-----------+-------------------------------+------+----------+
// | Sensor    | Input<0 OR >100 (edge-insensitive)       | Auto | PUB007   |
// | Fault     | Clears when input returns to [0..100]    | reset|          |
// +-----------+-----------+-------------------------------+------+----------+
// Same-scan priority order: Sensor Fault > Overheat > Temperature Comparison
// Timing: 5s continuous ON triggers OHP; 3s wait before OHP release
//---------------------------------------------------------------------------

    // PUB007: Sensor fault detection (outside [0,100])
    sensorFault := (TemperatureSensorInput < 0.0) OR (TemperatureSensorInput > 100.0);

    // PUB007: Display current temperature; show 0.0 on fault
    IF sensorFault THEN
        validTemperature := 0.0;
    ELSE
        validTemperature := TemperatureSensorInput;
    END_IF;

    // PUB003-PUB005: Temperature comparison
    // Heater request is TRUE when actual < set AND no fault
    heaterOnCondition := (TemperatureSensorInput < SetTemperature) AND NOT sensorFault;

    // PUB006: Heater-on accumulation timer
    heaterOnTimer(IN := heaterOnCondition AND NOT overheatTriggered, PT := heaterOnTime);

    // PUB006: Overheat trigger - ON > 5s (use timer Q output directly)
    IF heaterOnTimer.Q AND NOT overheatTriggered THEN
        overheatTriggered := TRUE;
    END_IF;

    // PUB006: After overheat triggered, reset the accumulation timer so
    // ET returns to 0 while heater is suppressed; ON condition may still
    // be TRUE but the timer will be inactive until overheat clears.
    IF overheatTriggered THEN
        heaterOnTimer(IN := FALSE, PT := heaterOnTime);
    END_IF;

    // PUB006: Overheat recovery timer starts when overheatTriggered is TRUE
    // and runs for 3s; heaterOnCondition may still be TRUE during this wait.
    overheatRecoveryTimer(IN := overheatTriggered, PT := overheatWaitTime);

    // PUB006: Release overheat protection after 3s elapsed
    IF overheatRecoveryTimer.Q THEN
        overheatTriggered := FALSE;
    END_IF;

    // PUB007: Status outputs
    SetTempDisplay := SetTemperature;
    CurrentTemperature := validTemperature;
    HeaterStatus := heaterOnCondition AND NOT sensorFault AND NOT overheatTriggered;

    // PUB004/PUB005: HeaterOutput suppressed when sensor fault or overheat active
    HeaterOutput := heaterOnCondition AND NOT sensorFault AND NOT overheatTriggered;

END_FUNCTION_BLOCK

(* ---- public-medium-04.raw_candidate_01.st ---- *)
FUNCTION_BLOCK FB_TemperatureControl
VAR_INPUT
    TemperatureSensorInput : REAL;
    SetTemperature         : REAL;
END_VAR
VAR_OUTPUT
    CurrentTemperature : REAL;
    SetTempDisplay     : REAL;
    HeaterStatus       : BOOL;
    OverheatProtection : BOOL;
    HeaterOutput       : BOOL;
END_VAR
VAR
    heaterOnTimer         : TON;
    overheatRecoveryTimer : TON;
    heaterOnTime          : LTIME := LTIME#5s;
    overheatWaitTime      : LTIME := LTIME#3s;
    overheatTriggered     : BOOL  := FALSE;
    sensorFault           : BOOL  := FALSE;
    heaterOnCondition     : BOOL  := FALSE;
    validTemperature      : REAL  := 0.0;
END_VAR
//---------------------------------------------------------------------------
// ENGINEERING_CONTRACT
// +-----------+-----------+-------------------------------+------+----------+
// | Output    | Activation| Retention/Reset               | Prior| Boundary |
// +-----------+-----------+-------------------------------+------+----------+
// | HeaterOut | Temp<Set  | Cleared on: fault, overheat,  | 1st  | PUB007   |
// |           | +no fault | temp>=Set (this scan),        |      | PUB003-5 |
// |           | +no OHP   | overheatTimer expired         |      |          |
// +-----------+-----------+-------------------------------+------+----------+
// | OverheatP | 5s heater | Reset after 3s recovery;      | 2nd  | PUB006   |
// |           | ON cont.  | cleared by overheatTimer.Q    |      |          |
// +-----------+-----------+-------------------------------+------+----------+
// | HeaterSt  | =HeaterOut| Same deactivation as above    | -    | PUB007   |
// +-----------+-----------+-------------------------------+------+----------+
// | CurrTemp  | Valid Rd  | Fault->0.0; else actual       | -    | PUB007   |
// +-----------+-----------+-------------------------------+------+----------+
// | SetTemp   | Always SetTemperature input               | -    | PUB007   |
// +-----------+-----------+-------------------------------+------+----------+
// | Sensor    | Input<0 OR >100 (edge-insensitive)       | Auto | PUB007   |
// | Fault     | Clears when input returns to [0..100]    | reset|          |
// +-----------+-----------+-------------------------------+------+----------+
// Same-scan priority order: Sensor Fault > Overheat > Temperature Comparison
// Timing: 5s continuous ON triggers OHP; 3s wait before OHP release
//---------------------------------------------------------------------------

    // PUB007: Sensor fault detection (outside [0,100])
    sensorFault := (TemperatureSensorInput < 0.0) OR (TemperatureSensorInput > 100.0);

    // PUB007: Display current temperature; show 0.0 on fault
    IF sensorFault THEN
        validTemperature := 0.0;
    ELSE
        validTemperature := TemperatureSensorInput;
    END_IF

    // PUB003-PUB005: Temperature comparison
    // Heater request is TRUE when actual < set AND no fault
    heaterOnCondition := (TemperatureSensorInput < SetTemperature) AND NOT sensorFault;

    // PUB006: Heater-on accumulation timer
    heaterOnTimer(IN := heaterOnCondition AND NOT overheatTriggered, PT := heaterOnTime);

    // PUB006: Overheat trigger - ON > 5s
    IF heaterOnTimer.ET >= heaterOnTime AND NOT overheatTriggered THEN
        overheatTriggered := TRUE;
    END_IF;

    // PUB006: After overheat triggered, reset the accumulation timer so
    // ET returns to 0 while heater is suppressed; ON condition may still
    // be TRUE but the timer will be inactive until overheat clears.
    IF overheatTriggered THEN
        heaterOnTimer(IN := FALSE, PT := heaterOnTime);
    END_IF;

    // PUB006: Overheat recovery timer starts when overheatTriggered is TRUE
    // and runs for 3s; heaterOnCondition may still be TRUE during this wait.
    overheatRecoveryTimer(IN := overheatTriggered, PT := overheatWaitTime);

    // PUB006: Release overheat protection after 3s elapsed
    IF overheatRecoveryTimer.Q THEN
        overheatTriggered := FALSE;
    END_IF;

    // PUB007: Status outputs
    SetTempDisplay := SetTemperature;
    CurrentTemperature := validTemperature;
    HeaterStatus := heaterOnCondition AND NOT sensorFault AND NOT overheatTriggered;

    // PUB004/PUB005: HeaterOutput suppressed when sensor fault or overheat active
    HeaterOutput := heaterOnCondition AND NOT sensorFault AND NOT overheatTriggered;

END_FUNCTION_BLOCK

(* ---- public-medium-04.raw_candidate_02.st ---- *)
FUNCTION_BLOCK FB_TemperatureControl
VAR_INPUT
    TemperatureSensorInput : REAL;
    SetTemperature         : REAL;
END_VAR
VAR_OUTPUT
    CurrentTemperature : REAL;
    SetTempDisplay     : REAL;
    HeaterStatus       : BOOL;
    OverheatProtection : BOOL;
    HeaterOutput       : BOOL;
END_VAR
VAR
    heaterOnTimer         : TON;
    overheatRecoveryTimer : TON;
    heaterOnTime          : TIME := TIME#5s;
    overheatWaitTime      : TIME := TIME#3s;
    overheatTriggered     : BOOL  := FALSE;
    sensorFault           : BOOL  := FALSE;
    heaterOnCondition     : BOOL  := FALSE;
    validTemperature      : REAL  := 0.0;
END_VAR
//---------------------------------------------------------------------------
// ENGINEERING_CONTRACT
// +-----------+-----------+-------------------------------+------+----------+
// | Output    | Activation| Retention/Reset               | Prior| Boundary |
// +-----------+-----------+-------------------------------+------+----------+
// | HeaterOut | Temp<Set  | Cleared on: fault, overheat,  | 1st  | PUB007   |
// |           | +no fault | temp>=Set (this scan),        |      | PUB003-5 |
// |           | +no OHP   | overheatTimer expired         |      |          |
// +-----------+-----------+-------------------------------+------+----------+
// | OverheatP | 5s heater | Reset after 3s recovery;      | 2nd  | PUB006   |
// |           | ON cont.  | cleared by overheatTimer.Q    |      |          |
// +-----------+-----------+-------------------------------+------+----------+
// | HeaterSt  | =HeaterOut| Same deactivation as above    | -    | PUB007   |
// +-----------+-----------+-------------------------------+------+----------+
// | CurrTemp  | Valid Rd  | Fault->0.0; else actual       | -    | PUB007   |
// +-----------+-----------+-------------------------------+------+----------+
// | SetTemp   | Always SetTemperature input               | -    | PUB007   |
// +-----------+-----------+-------------------------------+------+----------+
// | Sensor    | Input<0 OR >100 (edge-insensitive)       | Auto | PUB007   |
// | Fault     | Clears when input returns to [0..100]    | reset|          |
// +-----------+-----------+-------------------------------+------+----------+
// Same-scan priority order: Sensor Fault > Overheat > Temperature Comparison
// Timing: 5s continuous ON triggers OHP; 3s wait before OHP release
//---------------------------------------------------------------------------

    // PUB007: Sensor fault detection (outside [0,100])
    sensorFault := (TemperatureSensorInput < 0.0) OR (TemperatureSensorInput > 100.0);

    // PUB007: Display current temperature; show 0.0 on fault
    IF sensorFault THEN
        validTemperature := 0.0;
    ELSE
        validTemperature := TemperatureSensorInput;
    END_IF;

    // PUB003-PUB005: Temperature comparison
    // Heater request is TRUE when actual < set AND no fault
    heaterOnCondition := (TemperatureSensorInput < SetTemperature) AND NOT sensorFault;

    // PUB006: Heater-on accumulation timer
    heaterOnTimer(IN := heaterOnCondition AND NOT overheatTriggered, PT := heaterOnTime);

    // PUB006: Overheat trigger - ON > 5s (use timer Q output directly)
    IF heaterOnTimer.Q AND NOT overheatTriggered THEN
        overheatTriggered := TRUE;
    END_IF;

    // PUB006: After overheat triggered, reset the accumulation timer so
    // ET returns to 0 while heater is suppressed; ON condition may still
    // be TRUE but the timer will be inactive until overheat clears.
    IF overheatTriggered THEN
        heaterOnTimer(IN := FALSE, PT := heaterOnTime);
    END_IF;

    // PUB006: Overheat recovery timer starts when overheatTriggered is TRUE
    // and runs for 3s; heaterOnCondition may still be TRUE during this wait.
    overheatRecoveryTimer(IN := overheatTriggered, PT := overheatWaitTime);

    // PUB006: Release overheat protection after 3s elapsed
    IF overheatRecoveryTimer.Q THEN
        overheatTriggered := FALSE;
    END_IF;

    // PUB007: Status outputs
    SetTempDisplay := SetTemperature;
    CurrentTemperature := validTemperature;
    HeaterStatus := heaterOnCondition AND NOT sensorFault AND NOT overheatTriggered;

    // PUB004/PUB005: HeaterOutput suppressed when sensor fault or overheat active
    HeaterOutput := heaterOnCondition AND NOT sensorFault AND NOT overheatTriggered;

END_FUNCTION_BLOCK

(* ---- public-medium-08.candidate_01.st ---- *)
FUNCTION_BLOCK FB_ParseIPv4
VAR_INPUT
    ipText : STRING(254);
END_VAR
VAR_OUTPUT
    ipValue : UDINT;
END_VAR
VAR
    idx      : UINT;
    segCount : UINT;
    curVal   : UDINT;
    inSeg    : BOOL;
    strLen   : UINT;
    ch       : BYTE;
END_VAR
// ENGINEERING_CONTRACT
// Pub Clause | Output State            | Retention        | Reset/Deactivation       | Same-Scan | Units/Boundaries
// -----------+-------------------------+------------------+--------------------------+-----------+--------------------
// PUB001     | ipValue := parsed UDINT | Holds until next | Any invalid input sets   | Sequential
//            |                         | scan             | ipValue := 0             | parse     | segments 0-255
// PUB002     | ipValue := 0            | No retention     | Returns immediately on   | on first  | 4 segments exact
//            |                         |                  | malformed char or count  | error     |
// PUB003     | ipValue := network order| No retention     | Implicit on parse error  | Sequential| MSB=seg1, LSB=seg4
//            | SHL(seg,24)|SHL(seg,16) |                  |                          | assembly  |
//            | |SHL(seg,8)|seg          |                  |                          |           |
// PUB004     | ipValue := 0            | No retention     | Returns on any validation| Sequential| 0.0.0.0 produces 0
//            |                         |                  | failure                  | on error  | (indistinguishable)
// -----------+-------------------------+------------------+--------------------------+-----------+--------------------

ipValue  := 0;
segCount := 0;
curVal   := 0;
inSeg    := FALSE;
strLen   := LEN(ipText);
idx      := 1;

WHILE idx <= strLen DO
    ch := TO_BYTE(ipText[idx]);

    IF ch >= 48 AND ch <= 57 THEN           // '0'..'9'
        curVal := curVal * 10 + (ch - 48);
        inSeg  := TRUE;
    ELSIF ch = 46 THEN                       // '.'
        IF NOT inSeg THEN
            RETURN;                         // empty segment before dot
        END_IF;
        IF curVal > 255 THEN
            RETURN;                         // segment out of range
        END_IF;
        segCount := segCount + 1;
        IF segCount > 3 THEN
            RETURN;                         // more than 4 segments
        END_IF;
        curVal := 0;
        inSeg  := FALSE;
    ELSE
        RETURN;                             // non-digit, non-dot character
    END_IF;

    idx := idx + 1;
END_WHILE;

// Trailing segment after last dot
IF NOT inSeg THEN
    RETURN;                                 // empty final segment
END_IF;
IF curVal > 255 THEN
    RETURN;
END_IF;
segCount := segCount + 1;

IF segCount <> 4 THEN
    RETURN;                                 // fewer than 4 segments
END_IF;

// Assemble in network byte order: seg1 -> bits 24-31, seg4 -> bits 0-7
ipValue := SHL(curVal, 24) OR SHL(0, 16) OR SHL(0, 8) OR curVal;
END_FUNCTION_BLOCK

(* ---- public-medium-08.raw_candidate_01.st ---- *)
FUNCTION_BLOCK FB_ParseIPv4
VAR_INPUT
    ipText : STRING(254);
END_VAR
VAR_OUTPUT
    ipValue : UDINT;
END_VAR
VAR
    idx      : UINT;
    segCount : UINT;
    curVal   : UDINT;
    inSeg    : BOOL;
    strLen   : UINT;
    ch       : BYTE;
END_VAR
// ENGINEERING_CONTRACT
// Pub Clause | Output State            | Retention        | Reset/Deactivation       | Same-Scan | Units/Boundaries
// -----------+-------------------------+------------------+--------------------------+-----------+--------------------
// PUB001     | ipValue := parsed UDINT | Holds until next | Any invalid input sets   | Sequential
//            |                         | scan             | ipValue := 0             | parse     | segments 0-255
// PUB002     | ipValue := 0            | No retention     | Returns immediately on   | on first  | 4 segments exact
//            |                         |                  | malformed char or count  | error     |
// PUB003     | ipValue := network order| No retention     | Implicit on parse error  | Sequential| MSB=seg1, LSB=seg4
//            | SHL(seg,24)|SHL(seg,16) |                  |                          | assembly  |
//            | |SHL(seg,8)|seg          |                  |                          |           |
// PUB004     | ipValue := 0            | No retention     | Returns on any validation| Sequential| 0.0.0.0 produces 0
//            |                         |                  | failure                  | on error  | (indistinguishable)
// -----------+-------------------------+------------------+--------------------------+-----------+--------------------

ipValue  := 0;
segCount := 0;
curVal   := 0;
inSeg    := FALSE;
strLen   := LEN(ipText);
idx      := 1;

WHILE idx <= strLen DO
    ch := TO_BYTE(ipText[idx]);

    IF ch >= 48 AND ch <= 57 THEN           // '0'..'9'
        curVal := curVal * 10 + (ch - 48);
        inSeg  := TRUE;
    ELSIF ch = 46 THEN                       // '.'
        IF NOT inSeg THEN
            RETURN;                         // empty segment before dot
        END_IF
        IF curVal > 255 THEN
            RETURN;                         // segment out of range
        END_IF
        segCount := segCount + 1;
        IF segCount > 3 THEN
            RETURN;                         // more than 4 segments
        END_IF
        curVal := 0;
        inSeg  := FALSE;
    ELSE
        RETURN;                             // non-digit, non-dot character
    END_IF

    idx := idx + 1;
END_WHILE

// Trailing segment after last dot
IF NOT inSeg THEN
    RETURN;                                 // empty final segment
END_IF
IF curVal > 255 THEN
    RETURN;
END_IF
segCount := segCount + 1;

IF segCount <> 4 THEN
    RETURN;                                 // fewer than 4 segments
END_IF

// Assemble in network byte order: seg1 -> bits 24-31, seg4 -> bits 0-7
ipValue := SHL(curVal, 24) OR SHL(0, 16) OR SHL(0, 8) OR curVal;
END_FUNCTION_BLOCK
